FUNCTION_BLOCK FB_Recipe
VAR_INPUT
	pstRecipe				:POINTER TO ST_Recipe;
	bMemoRecipeUpdated		:BOOL:=FALSE;
	sRecipeDef				:STRING; (* current recipe definition *)
	bLoadDefault			:BOOL;
	sRecipesStoragePath		:STRING;
	bHMI_FrameActive		:BOOL;

END_VAR

VAR
	i						:INT;	
	RecipeManCommands 		:RecipeManCommands; (* Recipe Manager *)
	k						:INT;
	t1						:TON;
	check					:DWORD;
	INDEX					:INT:= 0;
	bReloadRecipes			:BOOL;
	rt_LoadDefault: R_TRIG;
	MessageBox			:MessageBox_Struct;
	arrLastReturn		: ARRAY[0..15] OF DWORD;
	LastReturn			:  DWORD;
	ton_RecipeUpdated: TON;
	sMessage: STRING;
	ton_SetStoragePath_Delay: TON;
	bSetStoragePath: BOOL:=TRUE;
	ton_SetStoragePathTimeOut: TON;
	bReturn: BOOL;
	
	ton_MessClear: TON;
	rt_Init: R_TRIG;
	sLastMessage: STRING;
	rt_Saved: R_TRIG;
	rt_FrameAvtive: R_TRIG;
	rt_LoadDefault1: R_TRIG;
END_VAR

act_SetStoragePath();
act_Disp();

IF pstRecipe^.bValidSelected THEN
	pstRecipe^.sSelectedReceipe:= pstRecipe^.arrRecipeNames[pstRecipe^.iRecipeIndex];
	pstRecipe^.bValidSelected:=FALSE;
END_IF

rt_FrameAvtive(CLK:=bHMI_FrameActive);
rt_LoadDefault1(CLK:=bLoadDefault);
IF pstRecipe^.bReInit OR rt_LoadDefault1.Q OR rt_FrameAvtive.Q THEN;
	pstRecipe^.bReInit:=FALSE;
	pstRecipe^.bInit:=FALSE;
	bSetStoragePath:=TRUE;
END_IF

t1(IN:=NOT pstRecipe^.bInit , PT:=T#0.5S);
IF (NOT pstRecipe^.bInit AND t1.Q) THEN
	
	IF NOT bSetStoragePath THEN;
		arrLastReturn[3]:=RecipeManCommands.ResetLastInfo();
		arrLastReturn[4]:=RecipeManCommands.ReloadRecipes(RecipeDefinitionName:=sRecipeDef);
		pstRecipe^.iRecipeCount:=RecipeManCommands.GetRecipeCount(sRecipeDef);
		FOR i := 0 TO GVL_Recipe.C_Max_RecipeFileNum DO
			pstRecipe^.arrRecipeNames[i] := '';
		END_FOR
		FOR i := 0 TO 1200 DO
			pstRecipe^.arrVariableNamesValue[i] := '';
			pstRecipe^.arrVariableValue[i] := '';
		END_FOR	
		(* save all recipe names of one recipe definition in an array *)
		arrLastReturn[0]:=RecipeManCommands.GetRecipeNames(sRecipeDef, ADR(pstRecipe^.arrRecipeNames),GVL_Recipe.C_Max_RecipeFileNum, 0);
		pstRecipe^.iRecipeIndex:=0;
		pstRecipe^.sLastSelectedReceipe:=pstRecipe^.sSelectedReceipe:=pstRecipe^.arrRecipeNames[0];
		pstRecipe^.bInit:=TRUE;
		pstRecipe^.bReInit:=FALSE;		
	END_IF

END_IF


rt_Init(CLK:=pstRecipe^.bInit);
IF pstRecipe^.bInit THEN

	IF pstRecipe^.sSelectedReceipe <> pstRecipe^.sLastSelectedReceipe 
	OR rt_Init.Q 
	OR rt_Saved.Q
	THEN;
				 
		arrLastReturn[1]:=RecipeManCommands.GetRecipeValues
			(
			RecipeDefinitionName:= sRecipeDef,
			RecipeName:= pstRecipe^.sSelectedReceipe, 
			pStrings:= ADR(pstRecipe^.arrVariableValue), 
			iSize:= 1200, 
			iStartIndex:= 0, 
			iStringLength:=80
			 );		
					
		arrLastReturn[2]:=RecipeManCommands.GetRecipeVariableNames
			(
			RecipeDefinitionName:=sRecipeDef,
			RecipeName:=pstRecipe^.sSelectedReceipe, 
			pStrings:= ADR(pstRecipe^.arrVariableNamesValue), 
			iSize:= 1200, 
			iStartIndex:= 0
			);
				
			pstRecipe^.bShowFile:=FALSE;
	END_IF
	pstRecipe^.sLastSelectedReceipe:=pstRecipe^.sSelectedReceipe;
END_IF


FOR i:=0 TO 15 DO
	IF arrLastReturn[i]<>0 THEN
		LastReturn:=arrLastReturn[i];
		EXIT;
	END_IF
	IF i=15 AND arrLastReturn[i]=0 THEN
		LastReturn:=0;
	END_IF
END_FOR

act_Cmd_List();

ACTION act_Cmd_List:
rt_LoadDefault(CLK:=bLoadDefault AND NOT bSetStoragePath);
IF rt_LoadDefault.Q THEN;
	pstRecipe^.sSelectedReceipe:='Default';
	pstRecipe^.bWriteToPLC_Cmd:=TRUE;
END_IF


IF pstRecipe^.bReloadRecipes THEN
	arrLastReturn[3]:=RecipeManCommands.ResetLastInfo();
	arrLastReturn[4]:=RecipeManCommands.ReloadRecipes(RecipeDefinitionName:=sRecipeDef);
	pstRecipe^.bReloadRecipes:=FALSE;
END_IF


IF pstRecipe^.bGetLastError THEN
	arrLastReturn[5]:=RecipeManCommands.GetLastError();
	pstRecipe^.bGetLastError:=FALSE;
END_IF


IF pstRecipe^.bResetLastError THEN
	arrLastReturn[6]:=RecipeManCommands.ResetLastError();
	pstRecipe^.bResetLastError:=FALSE;
	sMessage:='';
	FOR i:=0 TO 15 DO
		arrLastReturn[i]:=0;
	END_FOR	
END_IF

rt_Saved(CLK:=NOT pstRecipe^.bSaveFileCmd);
IF pstRecipe^.bSaveFileCmd  THEN
	sMessage:='cmd Save Recipe';
	IF  METH_Search(pstRecipe:=pstRecipe , sSearchRecipe:=pstRecipe^.sSelectedReceipe ) THEN
		//arrLastReturn[7]:=RecipeManCommands.ReadAndSaveRecipeAs(RecipeDefinitionName:=sRecipeDef,
		arrLastReturn[7]:=RecipeManCommands.ReadAndSaveRecipe(RecipeDefinitionName:=sRecipeDef,
			RecipeName:=pstRecipe^.sSelectedReceipe);// ,
			//FileName:='.txtrecipe' );
		sMessage:='cmd Save Recipe - Done';
		pstRecipe^.bSaveFileCmd:=FALSE;
	ELSE;
		sMessage:='cmd Save Recipe - Failed';
	END_IF
END_IF


IF pstRecipe^.bWriteToPLC_Cmd  THEN
	sMessage:='cmd Load Recipe';
	bMemoRecipeUpdated:=FALSE;
	IF  METH_Search(pstRecipe:=pstRecipe , sSearchRecipe:=pstRecipe^.sSelectedReceipe ) THEN
		arrLastReturn[8]:=RecipeManCommands.LoadRecipe(RecipeDefinitionName:= sRecipeDef, RecipeName:= pstRecipe^.sSelectedReceipe);
		arrLastReturn[9]:=RecipeManCommands.WriteRecipe(RecipeDefinitionName:= sRecipeDef, RecipeName:= pstRecipe^.sSelectedReceipe);
		sMessage:='cmd Load Recipe - Done';
		pstRecipe^.bWriteToPLC_Cmd:=FALSE;
		ton_RecipeUpdated.IN:=TRUE;
	ELSE;
		sMessage:='cmd Load Recipe - Failed';
	END_IF
END_IF
ton_RecipeUpdated(PT:=T#1S);
IF ton_RecipeUpdated.Q THEN;
	bMemoRecipeUpdated:=TRUE;	
	ton_RecipeUpdated.IN:=FALSE;
END_IF


IF pstRecipe^.bCreateRecipe AND pstRecipe^.sNewRecipeName <> '' THEN
	arrLastReturn[10]:=RecipeManCommands.CreateRecipe(sRecipeDef ,pstRecipe^.sNewRecipeName);
	sMessage:='cmd Create Recipe - Done';
	pstRecipe^.bCreateRecipe:=FALSE;
	pstRecipe^.bReInit:=TRUE;
END_IF


IF pstRecipe^.bDeleteRecipe THEN
	sMessage:='cmd Delete Recipe';
	IF  METH_Search(pstRecipe:=pstRecipe , sSearchRecipe:=pstRecipe^.sSelectedReceipe ) THEN
		arrLastReturn[11]:=RecipeManCommands.DeleteRecipe(sRecipeDef ,pstRecipe^.sSelectedReceipe);
		sMessage:='cmd Delete Recipe - Done';
		pstRecipe^.bDeleteRecipe:=FALSE;
		pstRecipe^.bReInit:=TRUE;
	ELSE;
		sMessage:='cmd Delete Recipe - Failed';
	END_IF
END_IF

ton_MessClear(PT:=T#30S);
IF sMessage<>sLastMessage THEN;
	ton_MessClear(IN:=FALSE);
	sLastMessage:=sMessage;
ELSIF sMessage<>'' THEN;
	ton_MessClear.IN:=TRUE;
ELSE;
	ton_MessClear.IN:=FALSE;
END_IF
IF ton_MessClear.Q THEN;
	sMessage:='';
END_IF
END_ACTION

ACTION act_Disp:

IF pstRecipe^.iDispSel<0 THEN; pstRecipe^.iDispSel:=0; END_IF
IF pstRecipe^.iDispSel>1180 THEN; pstRecipe^.iDispSel:=1180; END_IF

//FOR k:=iDispSel TO iDispSel+19 DO;
FOR k:=0 TO 20 DO;
	pstRecipe^.arrVariableDisp[0,k]:= INT_TO_STRING(pstRecipe^.iDispSel+k);
	pstRecipe^.arrVariableDisp[1,k]:=pstRecipe^.arrVariableNamesValue[pstRecipe^.iDispSel+k];
	pstRecipe^.arrVariableDisp[2,k]:=pstRecipe^.arrVariableValue[pstRecipe^.iDispSel+k];
END_FOR
END_ACTION

ACTION act_SetStoragePath:
ton_SetStoragePath_Delay(PT:=T#0.5S,IN:=bSetStoragePath);
ton_SetStoragePathTimeOut(PT:=T#2S);

IF ton_SetStoragePath_Delay.Q THEN;
	bReturn:=RecipeManCommands.SetStoragePath(stPath:=sRecipesStoragePath);
	//sMessage:='cmd Set Storage Path';
	IF bReturn THEN;
		bSetStoragePath:=FALSE;
		ton_SetStoragePathTimeOut.IN:=FALSE;
		//sMessage:='cmd Set Storage Path - Done';
	ELSE
		ton_SetStoragePathTimeOut.IN:=TRUE;
	END_IF
	
	IF ton_SetStoragePathTimeOut.Q THEN;
		bSetStoragePath:=FALSE;
		ton_SetStoragePathTimeOut.IN:=FALSE;
		//sMessage:='cmd Set Storage Path - Failed';		
	END_IF
END_IF
END_ACTION

METHOD METH_Search : BOOL
VAR_INPUT
	pstRecipe :POINTER TO ST_Recipe;
	sSearchRecipe	:STRING(30);
END_VAR

VAR
	i: INT;
END_VAR
METH_Search:=FALSE;
FOR i:= 0 TO GVL_Recipe.C_Max_RecipeFileNum DO
	IF sSearchRecipe = pstRecipe^.arrRecipeNames[i] THEN
		METH_Search:=TRUE;
		EXIT;
	END_IF
END_FOR
END_METHOD

END_FUNCTION_BLOCK

(* stored: Version 1.1.0.1, ProductVersion 3.1.4024.12
   POU FB_Recipe: Id {63aafca7-f761-4915-bd75-9a94b86d59ef}, SpecialFunc None
   Action act_Cmd_List: Id {6128ec74-fb63-4c1f-b6c7-01c4524738f9}
   Action act_Disp: Id {c0550086-68e6-4b05-93cc-ce9cbc221459}
   Action act_SetStoragePath: Id {69a5cd38-f127-4f75-bbaf-37404ec242ac}
   Method METH_Search: Id {007bd1bf-2c8b-4e7b-bd55-b9334aa3e650} *)
